Fanuc KAREL source: kd00057.KL

-- PROVISIONAL review KL for V940-1; original PC SHA256 7c1d4f304a3f2a1cd8a09c4d3e3a29c0d5f18555cf88797cba241264b36f478f
-- Incomplete behavior may be omitted. Consult companion uncertainty JSON. Do not deploy.
PROGRAM KD00057
%NOLOCKGROUP
VAR
  I : INTEGER
  J : INTEGER
  B : BOOLEAN
  R : REAL
  S : STRING[80]
-- UNRESOLVED_DECL P type=000101
-- UNRESOLVED_DECL Q type=000101
BEGIN
  -- V9_ZERO_TABLE_METADATA_HINT layout=0001; no indexed target words; source/name/runtime held
  -- UNRESOLVED_PC offsets 5-37; opcodes 01,22,1C,06,22,1C,07,82,0B
  -- UNRESOLVED_PC offsets 42-46; opcodes 7F
END KD00057
